(* IEC 61131-3 sources: repolevel_ST_code_completion/dataset/project_code/GreatExampleOfAdvantages/global, 1 file *)

(* ---- GVL_MQTT.st ---- *)
{attribute 'qualified_only'}
VAR_GLOBAL
	MQTT_IN_OUT:MQTT.MQTT_IN_OUT;
END_VAR
